Fanuc KAREL source: KO00142.KL

PROGRAM KO00142
%NOLOCKGROUP
VAR
  R: REAL
  CFG: CONFIG
  OUT: XYZWPR
  N: REAL
BEGIN
  N = 1
  R = 2.0
  CFG.CFG_FLIP = TRUE
  OUT = POS(R, R, R, N, R, R, CFG)
END KO00142
